(* IEC 61131-3 sources: PLC-Static-Analysis/modules/plc-rules/src/test/resources/PLCA-L003, 2 files *)

(* ---- compliant.st ---- *)
TYPE E_Color : (Red, Green); END_TYPE

PROGRAM P_L003ok
VAR
    n : INT;
    m : INT;
    r : REAL;
    b : BOOL;
    c : BOOL;
    q : BOOL;
    eColor : E_Color;
END_VAR
IF n < 10 THEN
    q := TRUE;
ELSIF n > 10 THEN
    q := FALSE;
ELSE
    b := TRUE;
END_IF
CASE eColor OF
    E_Color.Red: q := TRUE;
    E_Color.Green: q := FALSE;
ELSE
    b := TRUE;
END_CASE
IF r < 1.0 THEN
    q := TRUE;
ELSIF r > 1.0 THEN
    q := FALSE;
ELSE
    b := TRUE;
END_IF
END_PROGRAM

(* ---- noncompliant.st ---- *)
PROGRAM P_L003
VAR
    n : INT;
    m : INT;
    r : REAL;
    b : BOOL;
    c : BOOL;
    q : BOOL;
END_VAR
IF n < 10 THEN
    q := TRUE;
ELSIF n >= 10 THEN
    q := FALSE;
ELSE // PLCA-L003
    b := TRUE;
END_IF
IF b THEN
    q := TRUE;
ELSIF NOT b THEN
    q := FALSE;
ELSE // PLCA-L003
    c := TRUE;
END_IF
IF n > 0 THEN
    IF n > 5 THEN
        q := TRUE;
    ELSIF n <= 5 THEN
        q := FALSE;
    ELSE // PLCA-L003
        c := TRUE;
    END_IF
END_IF
END_PROGRAM
